(* IEC 61131-3 sources: POMIRTS_lab3/AS/Library/AsIODiag, 3 files *)

(* ---- AsIODiag.typ ---- *)
(********************************************************************
 * COPYRIGHT -- Bernecker + Rainer
 ********************************************************************
 * Library: AsIODiag
 * File: AsIODiag.typ
 * Author: B+R
 ********************************************************************
 * Data types of library AsIODiag
 ********************************************************************)

TYPE
END_TYPE

(* ---- AsIODiag.fun ---- *)
(********************************************************************
 * COPYRIGHT -- Bernecker + Rainer
 ********************************************************************
 * Library: AsIODiag
 * File: AsIODiag.fun
 * Author: B+R
 ********************************************************************
 * Functions and function blocks of library AsIODiag
 ********************************************************************)

FUNCTION_BLOCK DiagCreateInfo			(*collects information about the currently configured and/or inserted hardware modules; asynchronous execution*)
	VAR_INPUT
		enable       : BOOL; 			(*enables execution*)
		infoKind     : UDINT; 			(*type of information to be generated, e.g. asdiagPLUGGED, asdiagCONFIGURED, ..*)
	END_VAR

	VAR
        StateMan     : UINT;			(*internal variable*)
        ErrMan       : UINT;			(*internal variable*)
        Init         : UDINT;			(*internal variable*)
	END_VAR

	VAR_OUTPUT
		status       : UINT; 			(*execution status: ERR_OK, ERR_FUB_ENABLE_FALSE, ERR_FUB_BUSY, 0xXXXX = see help*)
        ident        : UDINT;			(*identifier of the generated information*)
        nrEntries    : UDINT;			(*number of generated information entries*)
	END_VAR
END_FUNCTION_BLOCK

FUNCTION_BLOCK DiagDisposeInfo			(*frees up the resources taken up by DiagCreateInfo(); asynchronous execution*)
	VAR_INPUT
		enable       : BOOL; 			(*enables execution*)
        ident        : UDINT;			(*identifier of the information to be freed up*)
	END_VAR

	VAR
        StateMan     : UINT;			(*internal variable*)
        ErrMan       : UINT;			(*internal variable*)
        Init         : UDINT;			(*internal variable*)
	END_VAR

	VAR_OUTPUT
		status  : UINT; 				(*execution status: ERR_OK, ERR_FUB_ENABLE_FALSE, ERR_FUB_BUSY, 0xXXXX = see help*)
	END_VAR
END_FUNCTION_BLOCK

FUNCTION_BLOCK DiagGetNumInfo			(*queries the numeric value of a specified information entry*)
	VAR_INPUT
		enable       : BOOL; 			(*enables execution*)
        ident        : UDINT;			(*identifier returned from DiagCreateInfo()*)
        index        : UDINT;			(*index of the entry [0..nrEntries-1]*)
        infoCode     : UDINT;			(*code of the desired information, e.g. asdiagMODUL_STATE, asdiagPLUGGED_MODNO, ..*)
	END_VAR

	VAR_OUTPUT
		status  : UINT; 				(*execution status: ERR_OK, ERR_FUB_ENABLE_FALSE, 0xXXXX = see help*)
        value   : UDINT;				(*numeric value*)
	END_VAR
END_FUNCTION_BLOCK

FUNCTION_BLOCK DiagGetStrInfo			(*queries the string value of a specified information entry*)
	VAR_INPUT
		enable       : BOOL; 			(*enables execution*)
        ident        : UDINT;			(*identifier returned from DiagCreateInfo()*)
        index        : UDINT;			(*index of the entry [0..nrEntries-1]*)
        infoCode     : UDINT;			(*code of the desired information*)
        pBuffer      : UDINT;			(*pointer to the return buffer*)
        bufferLen    : UDINT;			(*size of the return buffer*)
	END_VAR

	VAR_OUTPUT
		status   : UINT; 				(*execution status: ERR_OK, ERR_FUB_ENABLE_FALSE, 0xXXXX = see help*)
        stringLen: UDINT;				(*string length of the original data*)
	END_VAR
END_FUNCTION_BLOCK

(* ---- AsIODiag.var ---- *)
(********************************************************************
 * COPYRIGHT -- Bernecker + Rainer
 ********************************************************************
 * Library: AsIODiag
 * File: AsIODiag.var
 * Author: B+R
 ********************************************************************
 * Local variables of library AsIODiag
 ********************************************************************)

VAR CONSTANT

   asdiagERR_NOMEM  	: UINT := 30801; 		(*not enough memory to process the information*)
   asdiagERR_IDENT 	    : UINT := 30802; 		(*invalid ID*)
   asdiagERR_INDEX 	    : UINT := 30803; 		(*index out of range [0..nrEntries-1]*)
   asdiagERR_INFOCODE   : UINT := 30804; 		(*unknown infoCode parameter*)
   asdiagERR_INFOKIND   : UINT := 30805; 		(*unknown infoKind parameter*)

(* infoCode GetNumInfo *)
   asdiagMODUL_STATE  	: UDINT :=  1;			(*module state: 0x01 Module configured only, 0x02 Module inserted only, ..*)
   asdiagPLUGGED_MODNO 	: UDINT :=  2;			(*module code of inserted module*)
   asdiagCONFIG_MODNO 	: UDINT :=  3;			(*module code of configured module*)
   asdiagPLUGGED_FAMILY : UDINT :=	4;			(*family code of the inserted module*)
   asdiagCONFIG_FAMILY 	: UDINT :=  5;			(*family code of the configured module*)
   asdiagPLUGGED_USETYPE: UDINT := 	6;			(*use type of the inserted module*)
   asdiagCONFIG_USETYPE : UDINT :=	7; 			(*use type of the configured module*)
   asdiagSERIAL_NUMBER  : UDINT :=  8;          (*serial number of inserted module*)

(* infoCode GetStrInfo *)
   asdiagPATH  	        : UDINT :=	1001;		(*path of the module (e.g. "SL6.IF2.ST3.SL6.SS4"); the CPU path is "$root"*)
   asdiagPLUGGED_MODULE : UDINT :=	1002;		(*model number of the inserted module*)
   asdiagCONFIG_MODULE 	: UDINT :=	1003;		(*model number of the configured module*)
   asdiagPLUGGED_BUS 	: UDINT :=	1004;		(*bus system of the inserted module*)
   asdiagCONFIG_BUS 	: UDINT :=	1005;		(*bus system of the configured module*)
   asdiagHARDWARE_MODULE_NAME : UDINT := 1006;  (*hardware module name*)

(* infoKind *)
   asdiagPLUGGED  	: UDINT :=	1;				(*information about inserted modules*)
   asdiagCONFIGURED : UDINT :=	2;				(*information about configured modules*)
   asdiagALL 	    : UDINT :=	3;				(*information about inserted and configured modules*)
END_VAR
